FUNCTION F_CheckLowNibbleLEDState : BOOL
VAR_IN_OUT CONSTANT
    nValue: BYTE;
END_VAR
VAR_INPUT
    bFlashOn: BOOL;
END_VAR
VAR
    nNibble: BYTE;
END_VAR

nNibble := nValue AND BYTE#16#0F;
F_CheckLowNibbleLEDState := (nNibble <> BYTE#0) AND ((nNibble <> BYTE#3) OR bFlashOn);

END_FUNCTION

(* stored: Version 1.1.0.1
   POU F_CheckLowNibbleLEDState: Id {c6dd8d8f-cdc8-06f6-20dd-7f5d2737e40d}, SpecialFunc None *)
